// TIA Portal project "PLC_2_LINE2" (V18)

(* hardware
DEVICE "S7-1500/ET200MP station_1"  S7-1500 station
   slot 0: "Rail_0"  Rack  6ES7 590-1***0-0AA0
   slot 1: "PLC_2"  CPU 1511-1 PN  6ES7 511-1AK02-0AB0  V2.9
      slot 3: "CPU display_1"  6ES7591-1AA00-0AA0
      slot 32768: "PROFINET interface_1"  X1
         slot 32769: "Port_1"  X1 P1
         slot 32770: "Port_2"  X1 P2
      slot 34817: "Virtual CP interface port_1"  Virtual CP interface port  Virtual CP interface port
   slot 2: "DI 32x24VDC HF_1"  DI 32x24VDC HF  6ES7 521-1BL00-0AB0  V2.2
   slot 3: "DQ 32x24VDC/0.5A HF_1"  DQ 32x24VDC/0.5A HF  6ES7 522-1BL01-0AB0  V1.1
*)

// ===== PLC "PLC_2"  CPU 1511-1 PN =====

VAR_GLOBAL   // PLC tag table "Default tag table"
   "Tag_1" AT %I4.3 : Bool;
   "Tag_2" AT %I4.4 : Bool;
   "Tag_3" AT %I4.5 : Bool;
   "Tag_4" AT %I4.0 : Bool;
   "Tag_5" AT %I4.1 : Bool;
   "Tag_6" AT %I5.0 : Bool;
   "Tag_7" AT %I5.2 : Bool;
   "Tag_8" AT %I6.1 : Bool;
   "Tag_9" AT %I5.3 : Bool;
   "Tag_10" AT %I5.4 : Bool;
   "Tag_11" AT %I5.5 : Bool;
   "Tag_12" AT %I5.6 : Bool;
   "Tag_13" AT %I5.7 : Bool;
   "Tag_14" AT %I6.0 : Bool;
   "Tag_15" AT %Q1.6 : Bool;
   "Tag_16" AT %Q1.7 : Bool;
   "Tag_17" AT %Q2.0 : Bool;
   "Tag_18" AT %Q2.1 : Bool;
   "Tag_19" AT %Q2.2 : Bool;
   "Tag_20" AT %Q2.3 : Bool;
   "Tag_21" AT %I0.3 : Bool;
   "Tag_22" AT %I0.4 : Bool;
   "Tag_23" AT %I0.5 : Bool;
   "Tag_24" AT %I0.0 : Bool;
   "Tag_25" AT %I0.1 : Bool;
   "Tag_26" AT %I1.0 : Bool;
   "Tag_27" AT %I2.7 : Bool;
   "Tag_28" AT %I3.1 : Bool;
   "Tag_29" AT %I1.6 : Bool;
   "Tag_30" AT %I1.7 : Bool;
   "Tag_31" AT %I2.0 : Bool;
   "Tag_32" AT %I2.1 : Bool;
   "Tag_33" AT %I2.2 : Bool;
   "Tag_34" AT %I2.3 : Bool;
   "Tag_35" AT %I2.4 : Bool;
   "Tag_36" AT %I2.5 : Bool;
   "Tag_37" AT %I2.6 : Bool;
   "Tag_38" AT %I3.0 : Bool;
   "Tag_39" AT %Q0.4 : Bool;
   "Tag_40" AT %Q0.5 : Bool;
   "Tag_41" AT %Q0.6 : Bool;
   "Tag_42" AT %Q0.7 : Bool;
   "Tag_43" AT %Q1.0 : Bool;
   "Tag_44" AT %Q1.1 : Bool;
END_VAR

TYPE "typeTask"
   STRUCT
      station : Int;
      dwell_s : Int;
      crane : String[4];
      tank_name : String[10];
      prev : Int;
      next : Int;
      status : Int;
   END_STRUCT;
END_TYPE

TYPE "typeCraneData"
   STRUCT
      task_count : Int;
      tasks : Array[1..20] of "typeTask";
      cmd_send : Bool;
      sts_busy : Bool;
      sts_done : Bool;
      sts_step : Int;
      sts_state : Int;
      ls_at : Array[0..20] of Bool;
      ls_dip : Bool;
      ls_up : Bool;
      ls_mid : Bool;
      btn_start : Bool;
      mv_fwd : Bool;
      mv_rev : Bool;
      mv_up : Bool;
      mv_down : Bool;
      estop : Bool;
      auto : Bool;
      cmd_reset : Bool;
      cmd_stop : Bool;
      pos : Array[0..20] of Int;
   END_STRUCT;
END_TYPE

DATA_BLOCK "Crane2Data"   // DB1
{ S7_Optimized_Access := 'TRUE' }
VERSION : 0.1
BEGIN
   pos[0] := 8;
   pos[1] := 1;
   pos[2] := 2;
   pos[3] := 3;
   pos[4] := 4;
   pos[5] := 5;
   pos[6] := 6;
   pos[7] := 7;
END_DATA_BLOCK

DATA_BLOCK "Crane3Data"   // DB2
{ S7_Optimized_Access := 'TRUE' }
VERSION : 0.1
BEGIN
   pos[0] := 20;
   pos[1] := 19;
   pos[8] := 9;
   pos[9] := 10;
   pos[10] := 11;
   pos[11] := 12;
   pos[12] := 13;
   pos[13] := 14;
   pos[14] := 15;
   pos[15] := 16;
   pos[16] := 17;
   pos[17] := 18;
   pos[18] := 19;
END_DATA_BLOCK

DATA_BLOCK "Crane2_Seq_DB"   // DB3
{ S7_Optimized_Access := 'TRUE' }
VERSION : 0.1
// stored: InstanceOfName CraneSequencer
"CraneSequencer"
BEGIN
END_DATA_BLOCK

DATA_BLOCK "Crane3_Seq_DB"   // DB4
{ S7_Optimized_Access := 'TRUE' }
VERSION : 0.1
// stored: InstanceOfName CraneSequencer
"CraneSequencer"
BEGIN
END_DATA_BLOCK

FUNCTION_BLOCK "CraneSequencer"   // FB1, SCL
{ S7_Optimized_Access := 'TRUE' }
VERSION : 0.1
   VAR_IN_OUT
      d : "typeCraneData";
   END_VAR
   VAR
      state : Int;
      idx : Int;
      count : Int;
      cur : Int;
      prevSend : Bool;
      tHold : TON_TIME;
      tDwell : TON_TIME;
   END_VAR
   VAR_TEMP
      target : Int;
      arrived : Bool;
   END_VAR
BEGIN
   // ============================================================================
   //  CraneSequencer  —  GENERIC per-crane batch sequencer  (LIBRARY block)
   // ----------------------------------------------------------------------------
   //  ONE function block reused by EVERY crane on EVERY PLC. Call once per scan
   //  from OB1, passing that crane's data block as the InOut #d. No copy, no
   //  find/replace — the crane it drives is chosen entirely by which DB you pass.
   //
   //  Block type : FUNCTION BLOCK (FB), language SCL.
   //  InOut      : d : "typeCraneData"           // the whole crane interface (a DB of this UDT)
   //  Static     : state:Int, idx:Int, count:Int, cur:Int, prevSend:Bool,
   //               tHold:TON_TIME, tDwell:TON_TIME
   //  Temp       : target:Int, arrived:Bool
   //
   //  OB1 (per crane):  CraneSequencer(d := "Crane6Data")   // its own instance DB
   //                    CraneSequencer(d := "Crane7AData")
   //
   //  Stations: 0=Parking  1=Loading  2..N = tanks (tank number + 1).
   //  States : 0 IDLE · 10 GO_LOAD · 20 LOWER_LOAD · 30 WAIT_BTN · 40 LIFT_LOAD
   //           50 GO_TANK · 60 LOWER_TANK · 70 DWELL · 80 LIFT_TANK · 85 GO_PARK · 90 DONE
   //
   //  DIRECTION IS BY PHYSICAL POSITION, NOT STATION NUMBER.
   //  The plant is NOT laid out in station-number order: Parking sits WEST of Loading, and a
   //  downstream crane's Loading is a transfer tank at the far (West) end. So travel direction
   //  is decided from #d.pos[station] — the physical left→right position of each station
   //  (1 = East-most … larger = further West). TravelTo drives WEST (mv_fwd → R-West) toward a
   //  HIGHER pos, EAST (mv_rev → R-East) toward a LOWER pos. The station's arrival switch is still
   //  #d.ls_at[station]. **Set #d.pos[] per crane** — see the PLC's position-map doc.
   //
   //  COMMANDS (app/Manager writes these):
   //    cmd_send  — arm a batch (rising edge, from IDLE).
   //    cmd_stop  — EMERGENCY HOLD: kills all motion immediately, latches state 100 (STOPPED).
   //                Does NOT clear the recipe. Clear it (and Reset) to move again.
   //    cmd_reset — CLEAN/HOME: lift clear → travel to Parking → wipe the recipe → IDLE.
   //                "As if no recipe was sent, crane back at its home." PLC clears cmd_reset when done.
   //  Extra states: 100 STOPPED · 110 RESET_LIFT · 120 RESET_HOME.
   // ============================================================================

   // ---- command overrides (run BEFORE the state machine, highest priority) ----
   IF #d.cmd_stop THEN                       // immediate emergency hold (latched)
       #d.mv_fwd := FALSE;
       #d.mv_rev := FALSE;
       #d.mv_up := FALSE;
       #d.mv_down := FALSE;
       #d.sts_busy := FALSE;
       #state := 100;
   ELSIF #d.cmd_reset AND #state <> 110 AND #state <> 120 THEN   // start homing/clear (if not already)
       // Wipe the recipe IMMEDIATELY (visible at once), then home the crane.
       #d.task_count := 0;
       #d.sts_step := 0;
       #d.sts_done := FALSE;
       #d.cmd_send := FALSE;
       #idx := 0;
       #count := 0;
       #d.sts_busy := TRUE;
       #state := 110;
   END_IF;

   #d.sts_state := #state;

   CASE #state OF
       0:  // IDLE — parked, hoist up, motors off, waiting for a batch.
           #d.mv_fwd := FALSE;
           #d.mv_rev := FALSE;
           #d.mv_up := FALSE;
           #d.mv_down := FALSE;
           #d.sts_busy := FALSE;
           #d.sts_step := 0;
           IF #d.cmd_send AND NOT #prevSend AND #d.task_count > 0 THEN
               #count := #d.task_count;
               #idx := 1;
               #d.sts_done := FALSE;
               #d.sts_busy := TRUE;
               #state := 10;
           END_IF;

       10: // GO_LOAD — travel to the Loading Area (station 1).
           #d.sts_busy := TRUE;
           #target := 1;
           #arrived := "TravelTo"(target := #d.pos[#target], cur := #d.pos[#cur],
                                  atTarget := #d.ls_at[#target],
                                  fwd => #d.mv_fwd, rev => #d.mv_rev);
           IF #arrived THEN
               #cur := #target;
               #d.mv_fwd := FALSE;
               #d.mv_rev := FALSE;
               #state := 20;
           END_IF;

       20: // LOWER_LOAD — lower the hoist until the dip limit switch is made.
           #d.mv_up := FALSE;
           #d.mv_down := TRUE;
           IF #d.ls_dip THEN
               #d.mv_down := FALSE;
               #state := 30;
           END_IF;

       30: // WAIT_BTN — operator loads material, then HOLDS btn_start for 3 s.
           #tHold(IN := #d.btn_start,
                  PT := T#3S);
           IF #tHold.Q THEN
               #state := 40;
           END_IF;

       40: // LIFT_LOAD — raise the hoist clear before travelling.
           #d.mv_down := FALSE;
           #d.mv_up := TRUE;
           IF #d.ls_up THEN
               #d.mv_up := FALSE;
               #state := 50;
           END_IF;

       50: // GO_TANK — travel to THIS task's tank station (TravelTo reverses if lower).
           #d.sts_step := #idx;
           #d.tasks[#idx].status := 1;                  // running
           #target := #d.tasks[#idx].station;
           #arrived := "TravelTo"(target := #d.pos[#target], cur := #d.pos[#cur],
                                  atTarget := #d.ls_at[#target],
                                  fwd => #d.mv_fwd, rev => #d.mv_rev);
           IF #arrived THEN
               #cur := #target;
               #d.mv_fwd := FALSE;
               #d.mv_rev := FALSE;
               #state := 60;
           END_IF;

       60: // LOWER_TANK — dip into the tank until the dip limit switch is made.
           #d.mv_up := FALSE;
           #d.mv_down := TRUE;
           IF #d.ls_dip THEN
               #d.mv_down := FALSE;
               #state := 70;
           END_IF;

       70: // DWELL — hold in the tank for this task's dwell_s seconds.
           #tDwell(IN := TRUE,
                   PT := DINT_TO_TIME(INT_TO_DINT(#d.tasks[#idx].dwell_s) * 1000));
           IF #tDwell.Q THEN
               #tDwell(IN := FALSE,
                       PT := T#0S);        // reset the timer for the next tank
               #state := 80;
           END_IF;

       80: // LIFT_TANK — lift out, mark the task done, advance or finish.
           #d.mv_down := FALSE;
           #d.mv_up := TRUE;
           IF #d.ls_up THEN
               #d.mv_up := FALSE;
               #d.tasks[#idx].status := 2;              // done
               IF #idx < #count THEN
                   #idx := #idx + 1;
                   #state := 50;                        // next tank
               ELSE
                   #state := 85;                        // all tanks done
               END_IF;
           END_IF;

       85: // GO_PARK — return home to Parking (station 0).
           #target := 0;
           #arrived := "TravelTo"(target := #d.pos[#target], cur := #d.pos[#cur],
                                  atTarget := #d.ls_at[#target],
                                  fwd => #d.mv_fwd, rev => #d.mv_rev);
           IF #arrived THEN
               #cur := #target;
               #d.mv_fwd := FALSE;
               #d.mv_rev := FALSE;
               #state := 90;
           END_IF;

       90: // DONE — raise the done flag, wait for the app to acknowledge (cmd_send → FALSE).
           #d.sts_busy := FALSE;
           #d.sts_done := TRUE;
           IF NOT #d.cmd_send THEN
               #d.sts_done := FALSE;
               #d.sts_step := 0;
               #state := 0;
           END_IF;

       100: // STOPPED — emergency hold. Motors off; leaves only via Reset (cmd_reset).
           #d.mv_fwd := FALSE;
           #d.mv_rev := FALSE;
           #d.mv_up := FALSE;
           #d.mv_down := FALSE;
           #d.sts_busy := FALSE;

       110: // RESET_LIFT — raise the hoist clear before homing.
           #d.mv_down := FALSE;
           #d.mv_up := TRUE;
           IF #d.ls_up THEN
               #d.mv_up := FALSE;
               #state := 120;
           END_IF;

       120: // RESET_HOME — travel to Parking, then wipe the recipe → IDLE.
           #target := 0;
           #arrived := "TravelTo"(target := #d.pos[#target], cur := #d.pos[#cur],
                                  atTarget := #d.ls_at[#target],
                                  fwd => #d.mv_fwd, rev => #d.mv_rev);
           IF #arrived THEN
               #cur := 0;
               #d.mv_fwd := FALSE;
               #d.mv_rev := FALSE;
               #d.task_count := 0;          // "as if no recipe was sent"
               #d.sts_step := 0;
               #d.sts_done := FALSE;
               #d.sts_busy := FALSE;
               #d.cmd_send := FALSE;
               #d.cmd_reset := FALSE;      // handshake: reset complete
               #idx := 0;
               #count := 0;
               #state := 0;                 // IDLE
           END_IF;
   END_CASE;

   #prevSend := #d.cmd_send;   // edge memory (runs every scan, after the CASE)
END_FUNCTION_BLOCK

FUNCTION "IOMap" : Void   // FC1, SCL
{ S7_Optimized_Access := 'TRUE' }
VERSION : 0.1
BEGIN
   // ============================================================================
   //  IOMap  —  PLC_2 (Line 2, cranes 2 & 3)  —  real %I/%Q ↔ crane DB mirrors
   //  FUNCTION (FC), SCL, return Void, no params. Call FIRST in OB1.
   //  Addresses from docs/plc/plant-panel-layout.md (PLC_2). Station = tank.number + 1.
   //
   //  ROLES (confirmed from the plant picture, East→West):
   //    Crane 2 = ENTRY  — loads at LOAD (East end), runs 15-3…4-6A, parks P-2.
   //    Crane 3 = DOWNSTREAM — picks up at TRVL-2A (West), runs DRY-2A…4-6B, parks P-3.
   //  Direction is by physical position (see ./POSITION-MAP.md): mv_fwd=West, mv_rev=East.
   // ============================================================================

   // ============================ CRANE 2  (Crane2Data) — ENTRY crane ============
   //  Loads at the LOAD bay (station 1, physical East end). Tanks run West from there;
   //  Parking (P-2) sits West of its tanks.
   "Crane2Data".ls_mid := "Tag_1";      // LS_Mid_C2
   "Crane2Data".ls_up := "Tag_2";      // LS_Up_C2
   "Crane2Data".ls_dip := "Tag_3";      // LS_Down_C2
   "Crane2Data".estop := "Tag_4";      // E-Stop_SW_C2
   "Crane2Data".auto := "Tag_5";      // Auto_SW_C2
   "Crane2Data".btn_start := "Tag_6";      // UP_Pendant_C2
   "Crane2Data".ls_at[0] := "Tag_7";      // PRK-2A_C2  (Parking — station 0)
   "Crane2Data".ls_at[1] := "Tag_8";      // LOAD-2A_C2 (Loading — entry bay)  [VERIFY on Panel_2]
   "Crane2Data".ls_at[2] := "Tag_9";      // 15-3_C2   (tank 1 -> station 2)
   "Crane2Data".ls_at[3] := "Tag_10";      // 4-7_C2    (tank 2 -> station 3)
   "Crane2Data".ls_at[4] := "Tag_11";      // 4-9_C2    (tank 3 -> station 4)
   "Crane2Data".ls_at[5] := "Tag_12";      // INS-2A_C2 (tank 4 -> station 5)
   "Crane2Data".ls_at[6] := "Tag_13";      // 4-10_C2   (tank 5 -> station 6)
   "Crane2Data".ls_at[7] := "Tag_14";      // 4-6A_C2   (tank 6 -> station 7)
   "Tag_15" := "Crane2Data".mv_up;          // R-Up_C2
   "Tag_16" := "Crane2Data".mv_down;        // R-Down_C2
   "Tag_17" := "Crane2Data".mv_rev;         // R-East_C2   (East = reverse / lower position)
   "Tag_18" := "Crane2Data".mv_fwd;         // R-West_C2   (West = forward / higher position)
   "Tag_19" := "Crane2Data".mv_up OR "Crane2Data".mv_down;     // R-Hoist_C2
   "Tag_20" := "Crane2Data".mv_fwd OR "Crane2Data".mv_rev;     // R-Trolley_C2

   // ============================ CRANE 3  (Crane3Data) — DOWNSTREAM =============
   //  No LOAD bay — Loading (station 1) is the transfer pickup at TRVL-2A (West end),
   //  the same switch as station 18. Its tanks run East of TRVL-2A; Parking (P-3) is
   //  the West-most box.
   "Crane3Data".ls_mid := "Tag_21";      // LS_Mid_C3
   "Crane3Data".ls_up := "Tag_22";      // LS_Up_C3
   "Crane3Data".ls_dip := "Tag_23";      // LS_Down_C3
   "Crane3Data".estop := "Tag_24";      // E-Stop_SW_C3
   "Crane3Data".auto := "Tag_25";      // Auto_SW_C3
   "Crane3Data".btn_start := "Tag_26";      // UP_Pendant_C3
   "Crane3Data".ls_at[0] := "Tag_27";      // PRK-2B_C3  (Parking — station 0)
   "Crane3Data".ls_at[1] := "Tag_28";      // TRVL-2A_C3 (Loading = transfer pickup; same as station 18)
   "Crane3Data".ls_at[8] := "Tag_29";      // DRY-2A_C3 (tank 7  -> station 8)
   "Crane3Data".ls_at[9] := "Tag_30";      // 4-8_C3    (tank 8  -> station 9)
   "Crane3Data".ls_at[10] := "Tag_31";      // 4-1_C3    (tank 9  -> station 10)
   "Crane3Data".ls_at[11] := "Tag_32";      // 4-2_C3    (tank 10 -> station 11)
   "Crane3Data".ls_at[12] := "Tag_33";      // 4-3_C3    (tank 11 -> station 12)
   "Crane3Data".ls_at[13] := "Tag_34";      // 4-4_C3    (tank 12 -> station 13)
   "Crane3Data".ls_at[14] := "Tag_35";      // 4-5_C3    (tank 13 -> station 14)
   "Crane3Data".ls_at[15] := "Tag_36";      // INS-2B_C3 (tank 14 -> station 15)
   "Crane3Data".ls_at[16] := "Tag_37";      // 4-11_C3   (tank 15 -> station 16)
   "Crane3Data".ls_at[17] := "Tag_38";      // 4-6B_C3   (tank 16 -> station 17)
   "Crane3Data".ls_at[18] := "Tag_28";      // TRVL-2A_C3 (tank 17 -> station 18; = Loading pickup)
   "Tag_39" := "Crane3Data".mv_up;          // R-Up_C3
   "Tag_40" := "Crane3Data".mv_down;        // R-Down_C3
   "Tag_41" := "Crane3Data".mv_rev;         // R-East_C3
   "Tag_42" := "Crane3Data".mv_fwd;         // R-West_C3
   "Tag_43" := "Crane3Data".mv_up OR "Crane3Data".mv_down;     // R-Hoist_C3
   "Tag_44" := "Crane3Data".mv_fwd OR "Crane3Data".mv_rev;     // R-Trolley_C3
END_FUNCTION

FUNCTION "TravelTo" : Bool   // FC2, SCL
{ S7_Optimized_Access := 'TRUE' }
VERSION : 0.1
   VAR_INPUT
      target : Int;
      cur : Int;
      atTarget : Bool;
   END_VAR
   VAR_OUTPUT
      fwd : Bool;
      rev : Bool;
   END_VAR
BEGIN
   // TravelTo — pick the travel direction toward a target station.
   // Returns TRUE when the target limit switch is already made (arrived → stop).
   #fwd := FALSE;
   #rev := FALSE;

   IF #atTarget THEN
       ;                       // arrived: leave both motors off
   ELSIF #target > #cur THEN
       #fwd := TRUE;           // higher station number → travel forward
   ELSE
       #rev := TRUE;           // lower station number → travel reverse
   END_IF;

   #TravelTo := #atTarget;
END_FUNCTION

ORGANIZATION_BLOCK "Main"   // OB1, LAD, ProgramCycle
TITLE = "Main Program Sweep (Cycle)"
{ S7_Optimized_Access := 'TRUE' }
VERSION : 0.1
   VAR_INPUT
      Initial_Call : Bool;   // Initial call of this OB
      Remanence : Bool;   // =True, if remanent data are available
   END_VAR
BEGIN

REGION Network 1
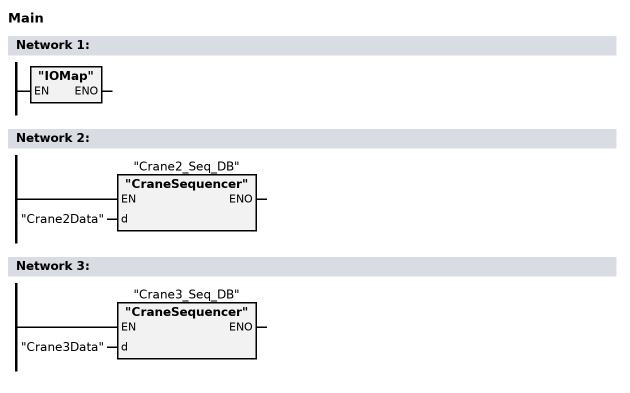
   RUNG wire#powerrail
      "IOMap"()
   END_RUNG
   // the same network as SCL:
   "IOMap"();
END_REGION

REGION Network 2
   RUNG wire#powerrail
      "Crane2_Seq_DB"(d := "Crane2Data")
   END_RUNG
   // the same network as SCL:
   "Crane2_Seq_DB"(d := "Crane2Data");   // "CraneSequencer"
END_REGION

REGION Network 3
   RUNG wire#powerrail
      "Crane3_Seq_DB"(d := "Crane3Data")
   END_RUNG
   // the same network as SCL:
   "Crane3_Seq_DB"(d := "Crane3Data");   // "CraneSequencer"
END_REGION
END_ORGANIZATION_BLOCK